// TIA Portal V19 export
// export: Created 2026-10-15T10:10:34.4181953Z, ExportSetting WithDefaults, DisplayName Totally Integrated Automation Portal, DisplayVersion V19, DisplayName TIA Portal Openness, DisplayVersion V19, DisplayName TIA Portal Version Control Interface, DisplayVersion V19, DisplayName STEP 7 Professional, DisplayVersion V19, DisplayName STEP 7 Safety, DisplayVersion V19, DisplayName WinCC Basic/Comfort/Advanced, DisplayVersion V19, DisplayName WinCC Unified, DisplayVersion V19
DATA_BLOCK "ROLL_HMI"   // DB3
{ S7_Optimized_Access := 'TRUE' }
VERSION : 0.1
// Flat, symbolic WinCC interface; TP900 control binding is a separate build step.
// stored: AutoNumber true, DBAccessibleFromOPCUA true, DBAccessibleFromWebserver true, IsOnlyStoredInLoadMemory false, IsRetainMemResEnabled false, IsWriteProtectedInAS false, MemoryReserve 100
   VAR
      Heartbeat : DInt;
      Connected : Bool;
      ManualFunction : Int := 255;
      GroundHeld : Bool;
      WorkHeld : Bool;
      KeyF : Array[1..16] of Bool;
      SelectedProgram : Int := 1;
      RecipeCommand : Int := 1;
      RecipeRequest : DInt;
      RecipeAck : DInt;
      RecipeError : Int;
      CurrentProgram : Int := 1;
      ParameterRequest : DInt;
      ParameterAck : DInt;
      ParameterDb : Int := 15;
      ParameterIndex : Int;
      ParameterValue : DInt;
      ParameterCurrentValue : DInt;
      ParameterSlotPresent : Bool;
      ParameterError : Int;
      Dwell1Seconds : Int := 360;
      Drain1Seconds : Int := 90;
      Ultrasound1 : Bool := TRUE;
      Dwell2Seconds : Int := 240;
      Drain2Seconds : Int := 60;
      Dwell3Seconds : Int := 300;
      Drain3Seconds : Int := 120;
      Dry4Seconds : Int := 400;
      BasketMotion : Int := 1;
      BathLift : Bool;
      ProcessTimer1Units : Int;
      ProcessTimer2Units : Int;
      StatusM : Array[0..255, 0..7] of Bool;
      LogicalOutputs : Array[16..25, 0..7] of Bool;
   END_VAR
BEGIN
END_DATA_BLOCK
